(* IEC 61131-3 sources: SemantiST/compiler/toolchain/compatibility/profiles/codesys-time, 1 file *)

(* ---- conversions.st ---- *)
(* Generated by compiler/toolchain/compatibility/profiles/generate_codesys.py
   from the pinned RuSTy standard library. Do not edit by hand.
   CODESYS TIME and TOD are 32-bit milliseconds, DATE and DT 32-bit seconds
   since 1970-01-01; RuSTy uses signed 64-bit nanoseconds. Adapters divide or
   multiply by the unit and keep the low bits on narrowing, as CODESYS does for
   integer conversions. TIME wrap-around at 2^32 ms is not simulated. *)

FUNCTION TIME_TO_BYTE : BYTE
VAR_INPUT IN : TIME; END_VAR
    TIME_TO_BYTE := LINT_TO_BYTE(TIME_TO_LINT(IN) / LINT#1000000);
END_FUNCTION

FUNCTION TIME_TO_WORD : WORD
VAR_INPUT IN : TIME; END_VAR
    TIME_TO_WORD := LINT_TO_WORD(TIME_TO_LINT(IN) / LINT#1000000);
END_FUNCTION

FUNCTION TIME_TO_DWORD : DWORD
VAR_INPUT IN : TIME; END_VAR
    TIME_TO_DWORD := LINT_TO_DWORD(TIME_TO_LINT(IN) / LINT#1000000);
END_FUNCTION

FUNCTION __CDS_TIME_TO_LWORD : LWORD
VAR_INPUT IN : TIME; END_VAR
    __CDS_TIME_TO_LWORD := LINT_TO_LWORD(TIME_TO_LINT(IN) / LINT#1000000);
END_FUNCTION

FUNCTION TIME_TO_SINT : SINT
VAR_INPUT IN : TIME; END_VAR
    TIME_TO_SINT := LINT_TO_SINT(TIME_TO_LINT(IN) / LINT#1000000);
END_FUNCTION

FUNCTION TIME_TO_USINT : USINT
VAR_INPUT IN : TIME; END_VAR
    TIME_TO_USINT := LINT_TO_USINT(TIME_TO_LINT(IN) / LINT#1000000);
END_FUNCTION

FUNCTION TIME_TO_INT : INT
VAR_INPUT IN : TIME; END_VAR
    TIME_TO_INT := LINT_TO_INT(TIME_TO_LINT(IN) / LINT#1000000);
END_FUNCTION

FUNCTION TIME_TO_UINT : UINT
VAR_INPUT IN : TIME; END_VAR
    TIME_TO_UINT := LINT_TO_UINT(TIME_TO_LINT(IN) / LINT#1000000);
END_FUNCTION

FUNCTION TIME_TO_DINT : DINT
VAR_INPUT IN : TIME; END_VAR
    TIME_TO_DINT := LINT_TO_DINT(TIME_TO_LINT(IN) / LINT#1000000);
END_FUNCTION

FUNCTION TIME_TO_UDINT : UDINT
VAR_INPUT IN : TIME; END_VAR
    TIME_TO_UDINT := LINT_TO_UDINT(TIME_TO_LINT(IN) / LINT#1000000);
END_FUNCTION

FUNCTION __CDS_TIME_TO_LINT : LINT
VAR_INPUT IN : TIME; END_VAR
    __CDS_TIME_TO_LINT := TIME_TO_LINT(IN) / LINT#1000000;
END_FUNCTION

FUNCTION __CDS_TIME_TO_ULINT : ULINT
VAR_INPUT IN : TIME; END_VAR
    __CDS_TIME_TO_ULINT := LINT_TO_ULINT(TIME_TO_LINT(IN) / LINT#1000000);
END_FUNCTION

FUNCTION TIME_TO_REAL : REAL
VAR_INPUT IN : TIME; END_VAR
    TIME_TO_REAL := LINT_TO_REAL(TIME_TO_LINT(IN) / LINT#1000000);
END_FUNCTION

FUNCTION __CDS_TIME_TO_LREAL : LREAL
VAR_INPUT IN : TIME; END_VAR
    __CDS_TIME_TO_LREAL := LINT_TO_LREAL(TIME_TO_LINT(IN) / LINT#1000000);
END_FUNCTION

FUNCTION TIME_TO_BOOL : BOOL
VAR_INPUT IN : TIME; END_VAR
    TIME_TO_BOOL := TIME_TO_LINT(IN) <> 0;
END_FUNCTION

FUNCTION BYTE_TO_TIME : TIME
VAR_INPUT IN : BYTE; END_VAR
VAR v : LINT; END_VAR
    v := IN;
    BYTE_TO_TIME := LINT_TO_TIME(v * LINT#1000000);
END_FUNCTION

FUNCTION WORD_TO_TIME : TIME
VAR_INPUT IN : WORD; END_VAR
VAR v : LINT; END_VAR
    v := IN;
    WORD_TO_TIME := LINT_TO_TIME(v * LINT#1000000);
END_FUNCTION

FUNCTION DWORD_TO_TIME : TIME
VAR_INPUT IN : DWORD; END_VAR
VAR v : LINT; END_VAR
    v := IN;
    DWORD_TO_TIME := LINT_TO_TIME(v * LINT#1000000);
END_FUNCTION

FUNCTION __CDS_LWORD_TO_TIME : TIME
VAR_INPUT IN : LWORD; END_VAR
VAR v : LINT; END_VAR
    v := IN;
    __CDS_LWORD_TO_TIME := LINT_TO_TIME(v * LINT#1000000);
END_FUNCTION

FUNCTION SINT_TO_TIME : TIME
VAR_INPUT IN : SINT; END_VAR
VAR v : LINT; END_VAR
    v := IN;
    SINT_TO_TIME := LINT_TO_TIME(v * LINT#1000000);
END_FUNCTION

FUNCTION USINT_TO_TIME : TIME
VAR_INPUT IN : USINT; END_VAR
VAR v : LINT; END_VAR
    v := IN;
    USINT_TO_TIME := LINT_TO_TIME(v * LINT#1000000);
END_FUNCTION

FUNCTION INT_TO_TIME : TIME
VAR_INPUT IN : INT; END_VAR
VAR v : LINT; END_VAR
    v := IN;
    INT_TO_TIME := LINT_TO_TIME(v * LINT#1000000);
END_FUNCTION

FUNCTION UINT_TO_TIME : TIME
VAR_INPUT IN : UINT; END_VAR
VAR v : LINT; END_VAR
    v := IN;
    UINT_TO_TIME := LINT_TO_TIME(v * LINT#1000000);
END_FUNCTION

FUNCTION DINT_TO_TIME : TIME
VAR_INPUT IN : DINT; END_VAR
VAR v : LINT; END_VAR
    v := IN;
    DINT_TO_TIME := LINT_TO_TIME(v * LINT#1000000);
END_FUNCTION

FUNCTION UDINT_TO_TIME : TIME
VAR_INPUT IN : UDINT; END_VAR
VAR v : LINT; END_VAR
    v := IN;
    UDINT_TO_TIME := LINT_TO_TIME(v * LINT#1000000);
END_FUNCTION

FUNCTION __CDS_LINT_TO_TIME : TIME
VAR_INPUT IN : LINT; END_VAR
VAR v : LINT; END_VAR
    v := IN;
    __CDS_LINT_TO_TIME := LINT_TO_TIME(v * LINT#1000000);
END_FUNCTION

FUNCTION __CDS_ULINT_TO_TIME : TIME
VAR_INPUT IN : ULINT; END_VAR
VAR v : LINT; END_VAR
    v := IN;
    __CDS_ULINT_TO_TIME := LINT_TO_TIME(v * LINT#1000000);
END_FUNCTION

FUNCTION REAL_TO_TIME : TIME
VAR_INPUT IN : REAL; END_VAR
VAR v : LINT; END_VAR
    v := REAL_TO_LINT(IN);
    REAL_TO_TIME := LINT_TO_TIME(v * LINT#1000000);
END_FUNCTION

FUNCTION __CDS_LREAL_TO_TIME : TIME
VAR_INPUT IN : LREAL; END_VAR
VAR v : LINT; END_VAR
    v := LREAL_TO_LINT(IN);
    __CDS_LREAL_TO_TIME := LINT_TO_TIME(v * LINT#1000000);
END_FUNCTION

FUNCTION BOOL_TO_TIME : TIME
VAR_INPUT IN : BOOL; END_VAR
    IF IN THEN
        BOOL_TO_TIME := LINT_TO_TIME(LINT#1000000);
    ELSE
        BOOL_TO_TIME := LINT_TO_TIME(LINT#0);
    END_IF;
END_FUNCTION

FUNCTION TOD_TO_BYTE : BYTE
VAR_INPUT IN : TIME_OF_DAY; END_VAR
    TOD_TO_BYTE := LINT_TO_BYTE(TOD_TO_LINT(IN) / LINT#1000000);
END_FUNCTION

FUNCTION TOD_TO_WORD : WORD
VAR_INPUT IN : TIME_OF_DAY; END_VAR
    TOD_TO_WORD := LINT_TO_WORD(TOD_TO_LINT(IN) / LINT#1000000);
END_FUNCTION

FUNCTION TOD_TO_DWORD : DWORD
VAR_INPUT IN : TIME_OF_DAY; END_VAR
    TOD_TO_DWORD := LINT_TO_DWORD(TOD_TO_LINT(IN) / LINT#1000000);
END_FUNCTION

FUNCTION __CDS_TOD_TO_LWORD : LWORD
VAR_INPUT IN : TIME_OF_DAY; END_VAR
    __CDS_TOD_TO_LWORD := LINT_TO_LWORD(TOD_TO_LINT(IN) / LINT#1000000);
END_FUNCTION

FUNCTION TOD_TO_SINT : SINT
VAR_INPUT IN : TIME_OF_DAY; END_VAR
    TOD_TO_SINT := LINT_TO_SINT(TOD_TO_LINT(IN) / LINT#1000000);
END_FUNCTION

FUNCTION TOD_TO_USINT : USINT
VAR_INPUT IN : TIME_OF_DAY; END_VAR
    TOD_TO_USINT := LINT_TO_USINT(TOD_TO_LINT(IN) / LINT#1000000);
END_FUNCTION

FUNCTION TOD_TO_INT : INT
VAR_INPUT IN : TIME_OF_DAY; END_VAR
    TOD_TO_INT := LINT_TO_INT(TOD_TO_LINT(IN) / LINT#1000000);
END_FUNCTION

FUNCTION TOD_TO_UINT : UINT
VAR_INPUT IN : TIME_OF_DAY; END_VAR
    TOD_TO_UINT := LINT_TO_UINT(TOD_TO_LINT(IN) / LINT#1000000);
END_FUNCTION

FUNCTION TOD_TO_DINT : DINT
VAR_INPUT IN : TIME_OF_DAY; END_VAR
    TOD_TO_DINT := LINT_TO_DINT(TOD_TO_LINT(IN) / LINT#1000000);
END_FUNCTION

FUNCTION TOD_TO_UDINT : UDINT
VAR_INPUT IN : TIME_OF_DAY; END_VAR
    TOD_TO_UDINT := LINT_TO_UDINT(TOD_TO_LINT(IN) / LINT#1000000);
END_FUNCTION

FUNCTION __CDS_TOD_TO_LINT : LINT
VAR_INPUT IN : TIME_OF_DAY; END_VAR
    __CDS_TOD_TO_LINT := TOD_TO_LINT(IN) / LINT#1000000;
END_FUNCTION

FUNCTION __CDS_TOD_TO_ULINT : ULINT
VAR_INPUT IN : TIME_OF_DAY; END_VAR
    __CDS_TOD_TO_ULINT := LINT_TO_ULINT(TOD_TO_LINT(IN) / LINT#1000000);
END_FUNCTION

FUNCTION TOD_TO_REAL : REAL
VAR_INPUT IN : TIME_OF_DAY; END_VAR
    TOD_TO_REAL := LINT_TO_REAL(TOD_TO_LINT(IN) / LINT#1000000);
END_FUNCTION

FUNCTION TOD_TO_LREAL : LREAL
VAR_INPUT IN : TIME_OF_DAY; END_VAR
    TOD_TO_LREAL := LINT_TO_LREAL(TOD_TO_LINT(IN) / LINT#1000000);
END_FUNCTION

FUNCTION TOD_TO_BOOL : BOOL
VAR_INPUT IN : TIME_OF_DAY; END_VAR
    TOD_TO_BOOL := TOD_TO_LINT(IN) <> 0;
END_FUNCTION

FUNCTION BYTE_TO_TOD : TIME_OF_DAY
VAR_INPUT IN : BYTE; END_VAR
VAR v : LINT; END_VAR
    v := IN;
    BYTE_TO_TOD := LINT_TO_TOD(v * LINT#1000000);
END_FUNCTION

FUNCTION WORD_TO_TOD : TIME_OF_DAY
VAR_INPUT IN : WORD; END_VAR
VAR v : LINT; END_VAR
    v := IN;
    WORD_TO_TOD := LINT_TO_TOD(v * LINT#1000000);
END_FUNCTION

FUNCTION DWORD_TO_TOD : TIME_OF_DAY
VAR_INPUT IN : DWORD; END_VAR
VAR v : LINT; END_VAR
    v := IN;
    DWORD_TO_TOD := LINT_TO_TOD(v * LINT#1000000);
END_FUNCTION

FUNCTION __CDS_LWORD_TO_TOD : TIME_OF_DAY
VAR_INPUT IN : LWORD; END_VAR
VAR v : LINT; END_VAR
    v := IN;
    __CDS_LWORD_TO_TOD := LINT_TO_TOD(v * LINT#1000000);
END_FUNCTION

FUNCTION SINT_TO_TOD : TIME_OF_DAY
VAR_INPUT IN : SINT; END_VAR
VAR v : LINT; END_VAR
    v := IN;
    SINT_TO_TOD := LINT_TO_TOD(v * LINT#1000000);
END_FUNCTION

FUNCTION USINT_TO_TOD : TIME_OF_DAY
VAR_INPUT IN : USINT; END_VAR
VAR v : LINT; END_VAR
    v := IN;
    USINT_TO_TOD := LINT_TO_TOD(v * LINT#1000000);
END_FUNCTION

FUNCTION INT_TO_TOD : TIME_OF_DAY
VAR_INPUT IN : INT; END_VAR
VAR v : LINT; END_VAR
    v := IN;
    INT_TO_TOD := LINT_TO_TOD(v * LINT#1000000);
END_FUNCTION

FUNCTION UINT_TO_TOD : TIME_OF_DAY
VAR_INPUT IN : UINT; END_VAR
VAR v : LINT; END_VAR
    v := IN;
    UINT_TO_TOD := LINT_TO_TOD(v * LINT#1000000);
END_FUNCTION

FUNCTION DINT_TO_TOD : TIME_OF_DAY
VAR_INPUT IN : DINT; END_VAR
VAR v : LINT; END_VAR
    v := IN;
    DINT_TO_TOD := LINT_TO_TOD(v * LINT#1000000);
END_FUNCTION

FUNCTION UDINT_TO_TOD : TIME_OF_DAY
VAR_INPUT IN : UDINT; END_VAR
VAR v : LINT; END_VAR
    v := IN;
    UDINT_TO_TOD := LINT_TO_TOD(v * LINT#1000000);
END_FUNCTION

FUNCTION __CDS_LINT_TO_TOD : TIME_OF_DAY
VAR_INPUT IN : LINT; END_VAR
VAR v : LINT; END_VAR
    v := IN;
    __CDS_LINT_TO_TOD := LINT_TO_TOD(v * LINT#1000000);
END_FUNCTION

FUNCTION __CDS_ULINT_TO_TOD : TIME_OF_DAY
VAR_INPUT IN : ULINT; END_VAR
VAR v : LINT; END_VAR
    v := IN;
    __CDS_ULINT_TO_TOD := LINT_TO_TOD(v * LINT#1000000);
END_FUNCTION

FUNCTION REAL_TO_TOD : TIME_OF_DAY
VAR_INPUT IN : REAL; END_VAR
VAR v : LINT; END_VAR
    v := REAL_TO_LINT(IN);
    REAL_TO_TOD := LINT_TO_TOD(v * LINT#1000000);
END_FUNCTION

FUNCTION LREAL_TO_TOD : TIME_OF_DAY
VAR_INPUT IN : LREAL; END_VAR
VAR v : LINT; END_VAR
    v := LREAL_TO_LINT(IN);
    LREAL_TO_TOD := LINT_TO_TOD(v * LINT#1000000);
END_FUNCTION

FUNCTION BOOL_TO_TOD : TIME_OF_DAY
VAR_INPUT IN : BOOL; END_VAR
    IF IN THEN
        BOOL_TO_TOD := LINT_TO_TOD(LINT#1000000);
    ELSE
        BOOL_TO_TOD := LINT_TO_TOD(LINT#0);
    END_IF;
END_FUNCTION

FUNCTION DATE_TO_BYTE : BYTE
VAR_INPUT IN : DATE; END_VAR
    DATE_TO_BYTE := LINT_TO_BYTE(DATE_TO_LINT(IN) / LINT#1000000000);
END_FUNCTION

FUNCTION DATE_TO_WORD : WORD
VAR_INPUT IN : DATE; END_VAR
    DATE_TO_WORD := LINT_TO_WORD(DATE_TO_LINT(IN) / LINT#1000000000);
END_FUNCTION

FUNCTION DATE_TO_DWORD : DWORD
VAR_INPUT IN : DATE; END_VAR
    DATE_TO_DWORD := LINT_TO_DWORD(DATE_TO_LINT(IN) / LINT#1000000000);
END_FUNCTION

FUNCTION __CDS_DATE_TO_LWORD : LWORD
VAR_INPUT IN : DATE; END_VAR
    __CDS_DATE_TO_LWORD := LINT_TO_LWORD(DATE_TO_LINT(IN) / LINT#1000000000);
END_FUNCTION

FUNCTION DATE_TO_SINT : SINT
VAR_INPUT IN : DATE; END_VAR
    DATE_TO_SINT := LINT_TO_SINT(DATE_TO_LINT(IN) / LINT#1000000000);
END_FUNCTION

FUNCTION DATE_TO_USINT : USINT
VAR_INPUT IN : DATE; END_VAR
    DATE_TO_USINT := LINT_TO_USINT(DATE_TO_LINT(IN) / LINT#1000000000);
END_FUNCTION

FUNCTION DATE_TO_INT : INT
VAR_INPUT IN : DATE; END_VAR
    DATE_TO_INT := LINT_TO_INT(DATE_TO_LINT(IN) / LINT#1000000000);
END_FUNCTION

FUNCTION DATE_TO_UINT : UINT
VAR_INPUT IN : DATE; END_VAR
    DATE_TO_UINT := LINT_TO_UINT(DATE_TO_LINT(IN) / LINT#1000000000);
END_FUNCTION

FUNCTION DATE_TO_DINT : DINT
VAR_INPUT IN : DATE; END_VAR
    DATE_TO_DINT := LINT_TO_DINT(DATE_TO_LINT(IN) / LINT#1000000000);
END_FUNCTION

FUNCTION DATE_TO_UDINT : UDINT
VAR_INPUT IN : DATE; END_VAR
    DATE_TO_UDINT := LINT_TO_UDINT(DATE_TO_LINT(IN) / LINT#1000000000);
END_FUNCTION

FUNCTION __CDS_DATE_TO_LINT : LINT
VAR_INPUT IN : DATE; END_VAR
    __CDS_DATE_TO_LINT := DATE_TO_LINT(IN) / LINT#1000000000;
END_FUNCTION

FUNCTION __CDS_DATE_TO_ULINT : ULINT
VAR_INPUT IN : DATE; END_VAR
    __CDS_DATE_TO_ULINT := LINT_TO_ULINT(DATE_TO_LINT(IN) / LINT#1000000000);
END_FUNCTION

FUNCTION DATE_TO_REAL : REAL
VAR_INPUT IN : DATE; END_VAR
    DATE_TO_REAL := LINT_TO_REAL(DATE_TO_LINT(IN) / LINT#1000000000);
END_FUNCTION

FUNCTION DATE_TO_LREAL : LREAL
VAR_INPUT IN : DATE; END_VAR
    DATE_TO_LREAL := LINT_TO_LREAL(DATE_TO_LINT(IN) / LINT#1000000000);
END_FUNCTION

FUNCTION DATE_TO_BOOL : BOOL
VAR_INPUT IN : DATE; END_VAR
    DATE_TO_BOOL := DATE_TO_LINT(IN) <> 0;
END_FUNCTION

FUNCTION BYTE_TO_DATE : DATE
VAR_INPUT IN : BYTE; END_VAR
VAR v : LINT; END_VAR
    v := IN;
    BYTE_TO_DATE := LINT_TO_DATE(v * LINT#1000000000);
END_FUNCTION

FUNCTION WORD_TO_DATE : DATE
VAR_INPUT IN : WORD; END_VAR
VAR v : LINT; END_VAR
    v := IN;
    WORD_TO_DATE := LINT_TO_DATE(v * LINT#1000000000);
END_FUNCTION

FUNCTION DWORD_TO_DATE : DATE
VAR_INPUT IN : DWORD; END_VAR
VAR v : LINT; END_VAR
    v := IN;
    DWORD_TO_DATE := LINT_TO_DATE(v * LINT#1000000000);
END_FUNCTION

FUNCTION __CDS_LWORD_TO_DATE : DATE
VAR_INPUT IN : LWORD; END_VAR
VAR v : LINT; END_VAR
    v := IN;
    __CDS_LWORD_TO_DATE := LINT_TO_DATE(v * LINT#1000000000);
END_FUNCTION

FUNCTION SINT_TO_DATE : DATE
VAR_INPUT IN : SINT; END_VAR
VAR v : LINT; END_VAR
    v := IN;
    SINT_TO_DATE := LINT_TO_DATE(v * LINT#1000000000);
END_FUNCTION

FUNCTION USINT_TO_DATE : DATE
VAR_INPUT IN : USINT; END_VAR
VAR v : LINT; END_VAR
    v := IN;
    USINT_TO_DATE := LINT_TO_DATE(v * LINT#1000000000);
END_FUNCTION

FUNCTION INT_TO_DATE : DATE
VAR_INPUT IN : INT; END_VAR
VAR v : LINT; END_VAR
    v := IN;
    INT_TO_DATE := LINT_TO_DATE(v * LINT#1000000000);
END_FUNCTION

FUNCTION UINT_TO_DATE : DATE
VAR_INPUT IN : UINT; END_VAR
VAR v : LINT; END_VAR
    v := IN;
    UINT_TO_DATE := LINT_TO_DATE(v * LINT#1000000000);
END_FUNCTION

FUNCTION DINT_TO_DATE : DATE
VAR_INPUT IN : DINT; END_VAR
VAR v : LINT; END_VAR
    v := IN;
    DINT_TO_DATE := LINT_TO_DATE(v * LINT#1000000000);
END_FUNCTION

FUNCTION UDINT_TO_DATE : DATE
VAR_INPUT IN : UDINT; END_VAR
VAR v : LINT; END_VAR
    v := IN;
    UDINT_TO_DATE := LINT_TO_DATE(v * LINT#1000000000);
END_FUNCTION

FUNCTION __CDS_LINT_TO_DATE : DATE
VAR_INPUT IN : LINT; END_VAR
VAR v : LINT; END_VAR
    v := IN;
    __CDS_LINT_TO_DATE := LINT_TO_DATE(v * LINT#1000000000);
END_FUNCTION

FUNCTION __CDS_ULINT_TO_DATE : DATE
VAR_INPUT IN : ULINT; END_VAR
VAR v : LINT; END_VAR
    v := IN;
    __CDS_ULINT_TO_DATE := LINT_TO_DATE(v * LINT#1000000000);
END_FUNCTION

FUNCTION REAL_TO_DATE : DATE
VAR_INPUT IN : REAL; END_VAR
VAR v : LINT; END_VAR
    v := REAL_TO_LINT(IN);
    REAL_TO_DATE := LINT_TO_DATE(v * LINT#1000000000);
END_FUNCTION

FUNCTION LREAL_TO_DATE : DATE
VAR_INPUT IN : LREAL; END_VAR
VAR v : LINT; END_VAR
    v := LREAL_TO_LINT(IN);
    LREAL_TO_DATE := LINT_TO_DATE(v * LINT#1000000000);
END_FUNCTION

FUNCTION BOOL_TO_DATE : DATE
VAR_INPUT IN : BOOL; END_VAR
    IF IN THEN
        BOOL_TO_DATE := LINT_TO_DATE(LINT#1000000000);
    ELSE
        BOOL_TO_DATE := LINT_TO_DATE(LINT#0);
    END_IF;
END_FUNCTION

FUNCTION DT_TO_BYTE : BYTE
VAR_INPUT IN : DATE_AND_TIME; END_VAR
    DT_TO_BYTE := LINT_TO_BYTE(DT_TO_LINT(IN) / LINT#1000000000);
END_FUNCTION

FUNCTION DT_TO_WORD : WORD
VAR_INPUT IN : DATE_AND_TIME; END_VAR
    DT_TO_WORD := LINT_TO_WORD(DT_TO_LINT(IN) / LINT#1000000000);
END_FUNCTION

FUNCTION DT_TO_DWORD : DWORD
VAR_INPUT IN : DATE_AND_TIME; END_VAR
    DT_TO_DWORD := LINT_TO_DWORD(DT_TO_LINT(IN) / LINT#1000000000);
END_FUNCTION

FUNCTION __CDS_DT_TO_LWORD : LWORD
VAR_INPUT IN : DATE_AND_TIME; END_VAR
    __CDS_DT_TO_LWORD := LINT_TO_LWORD(DT_TO_LINT(IN) / LINT#1000000000);
END_FUNCTION

FUNCTION DT_TO_SINT : SINT
VAR_INPUT IN : DATE_AND_TIME; END_VAR
    DT_TO_SINT := LINT_TO_SINT(DT_TO_LINT(IN) / LINT#1000000000);
END_FUNCTION

FUNCTION DT_TO_USINT : USINT
VAR_INPUT IN : DATE_AND_TIME; END_VAR
    DT_TO_USINT := LINT_TO_USINT(DT_TO_LINT(IN) / LINT#1000000000);
END_FUNCTION

FUNCTION DT_TO_INT : INT
VAR_INPUT IN : DATE_AND_TIME; END_VAR
    DT_TO_INT := LINT_TO_INT(DT_TO_LINT(IN) / LINT#1000000000);
END_FUNCTION

FUNCTION DT_TO_UINT : UINT
VAR_INPUT IN : DATE_AND_TIME; END_VAR
    DT_TO_UINT := LINT_TO_UINT(DT_TO_LINT(IN) / LINT#1000000000);
END_FUNCTION

FUNCTION DT_TO_DINT : DINT
VAR_INPUT IN : DATE_AND_TIME; END_VAR
    DT_TO_DINT := LINT_TO_DINT(DT_TO_LINT(IN) / LINT#1000000000);
END_FUNCTION

FUNCTION DT_TO_UDINT : UDINT
VAR_INPUT IN : DATE_AND_TIME; END_VAR
    DT_TO_UDINT := LINT_TO_UDINT(DT_TO_LINT(IN) / LINT#1000000000);
END_FUNCTION

FUNCTION __CDS_DT_TO_LINT : LINT
VAR_INPUT IN : DATE_AND_TIME; END_VAR
    __CDS_DT_TO_LINT := DT_TO_LINT(IN) / LINT#1000000000;
END_FUNCTION

FUNCTION __CDS_DT_TO_ULINT : ULINT
VAR_INPUT IN : DATE_AND_TIME; END_VAR
    __CDS_DT_TO_ULINT := LINT_TO_ULINT(DT_TO_LINT(IN) / LINT#1000000000);
END_FUNCTION

FUNCTION DT_TO_REAL : REAL
VAR_INPUT IN : DATE_AND_TIME; END_VAR
    DT_TO_REAL := LINT_TO_REAL(DT_TO_LINT(IN) / LINT#1000000000);
END_FUNCTION

FUNCTION DT_TO_LREAL : LREAL
VAR_INPUT IN : DATE_AND_TIME; END_VAR
    DT_TO_LREAL := LINT_TO_LREAL(DT_TO_LINT(IN) / LINT#1000000000);
END_FUNCTION

FUNCTION DT_TO_BOOL : BOOL
VAR_INPUT IN : DATE_AND_TIME; END_VAR
    DT_TO_BOOL := DT_TO_LINT(IN) <> 0;
END_FUNCTION

FUNCTION BYTE_TO_DT : DATE_AND_TIME
VAR_INPUT IN : BYTE; END_VAR
VAR v : LINT; END_VAR
    v := IN;
    BYTE_TO_DT := ULINT_TO_DT(LINT_TO_ULINT(v * LINT#1000000000));
END_FUNCTION

FUNCTION WORD_TO_DT : DATE_AND_TIME
VAR_INPUT IN : WORD; END_VAR
VAR v : LINT; END_VAR
    v := IN;
    WORD_TO_DT := ULINT_TO_DT(LINT_TO_ULINT(v * LINT#1000000000));
END_FUNCTION

FUNCTION DWORD_TO_DT : DATE_AND_TIME
VAR_INPUT IN : DWORD; END_VAR
VAR v : LINT; END_VAR
    v := IN;
    DWORD_TO_DT := ULINT_TO_DT(LINT_TO_ULINT(v * LINT#1000000000));
END_FUNCTION

FUNCTION __CDS_LWORD_TO_DT : DATE_AND_TIME
VAR_INPUT IN : LWORD; END_VAR
VAR v : LINT; END_VAR
    v := IN;
    __CDS_LWORD_TO_DT := ULINT_TO_DT(LINT_TO_ULINT(v * LINT#1000000000));
END_FUNCTION

FUNCTION SINT_TO_DT : DATE_AND_TIME
VAR_INPUT IN : SINT; END_VAR
VAR v : LINT; END_VAR
    v := IN;
    SINT_TO_DT := ULINT_TO_DT(LINT_TO_ULINT(v * LINT#1000000000));
END_FUNCTION

FUNCTION USINT_TO_DT : DATE_AND_TIME
VAR_INPUT IN : USINT; END_VAR
VAR v : LINT; END_VAR
    v := IN;
    USINT_TO_DT := ULINT_TO_DT(LINT_TO_ULINT(v * LINT#1000000000));
END_FUNCTION

FUNCTION INT_TO_DT : DATE_AND_TIME
VAR_INPUT IN : INT; END_VAR
VAR v : LINT; END_VAR
    v := IN;
    INT_TO_DT := ULINT_TO_DT(LINT_TO_ULINT(v * LINT#1000000000));
END_FUNCTION

FUNCTION UINT_TO_DT : DATE_AND_TIME
VAR_INPUT IN : UINT; END_VAR
VAR v : LINT; END_VAR
    v := IN;
    UINT_TO_DT := ULINT_TO_DT(LINT_TO_ULINT(v * LINT#1000000000));
END_FUNCTION

FUNCTION DINT_TO_DT : DATE_AND_TIME
VAR_INPUT IN : DINT; END_VAR
VAR v : LINT; END_VAR
    v := IN;
    DINT_TO_DT := ULINT_TO_DT(LINT_TO_ULINT(v * LINT#1000000000));
END_FUNCTION

FUNCTION UDINT_TO_DT : DATE_AND_TIME
VAR_INPUT IN : UDINT; END_VAR
VAR v : LINT; END_VAR
    v := IN;
    UDINT_TO_DT := ULINT_TO_DT(LINT_TO_ULINT(v * LINT#1000000000));
END_FUNCTION

FUNCTION LINT_TO_DT : DATE_AND_TIME
VAR_INPUT IN : LINT; END_VAR
VAR v : LINT; END_VAR
    v := IN;
    LINT_TO_DT := ULINT_TO_DT(LINT_TO_ULINT(v * LINT#1000000000));
END_FUNCTION

FUNCTION __CDS_ULINT_TO_DT : DATE_AND_TIME
VAR_INPUT IN : ULINT; END_VAR
VAR v : LINT; END_VAR
    v := IN;
    __CDS_ULINT_TO_DT := ULINT_TO_DT(LINT_TO_ULINT(v * LINT#1000000000));
END_FUNCTION

FUNCTION REAL_TO_DT : DATE_AND_TIME
VAR_INPUT IN : REAL; END_VAR
VAR v : LINT; END_VAR
    v := REAL_TO_LINT(IN);
    REAL_TO_DT := ULINT_TO_DT(LINT_TO_ULINT(v * LINT#1000000000));
END_FUNCTION

FUNCTION LREAL_TO_DT : DATE_AND_TIME
VAR_INPUT IN : LREAL; END_VAR
VAR v : LINT; END_VAR
    v := LREAL_TO_LINT(IN);
    LREAL_TO_DT := ULINT_TO_DT(LINT_TO_ULINT(v * LINT#1000000000));
END_FUNCTION

FUNCTION BOOL_TO_DT : DATE_AND_TIME
VAR_INPUT IN : BOOL; END_VAR
    IF IN THEN
        BOOL_TO_DT := ULINT_TO_DT(LINT_TO_ULINT(LINT#1000000000));
    ELSE
        BOOL_TO_DT := ULINT_TO_DT(LINT_TO_ULINT(LINT#0));
    END_IF;
END_FUNCTION

FUNCTION TOD_TO_TIME : TIME
VAR_INPUT IN : TIME_OF_DAY; END_VAR
    TOD_TO_TIME := LINT_TO_TIME(TOD_TO_LINT(IN));
END_FUNCTION

FUNCTION TIME_TO_TOD : TIME_OF_DAY
VAR_INPUT IN : TIME; END_VAR
    TIME_TO_TOD := LINT_TO_TOD(TIME_TO_LINT(IN));
END_FUNCTION

FUNCTION DATE_TO_DT : DATE_AND_TIME
VAR_INPUT IN : DATE; END_VAR
    DATE_TO_DT := ULINT_TO_DT(LINT_TO_ULINT(DATE_TO_LINT(IN)));
END_FUNCTION
